TYPE ST_CamStatus :
STRUCT
    eState : E_CamMachineState;
    eProcessPhase : E_CamProcessPhase;
    bPowerEnabled : BOOL;
    bReferenced : BOOL;
    bRecipeLoaded : BOOL;
    bCamActive : BOOL;
    bRunning : BOOL;
    bBusy : BOOL;
    eApplicationError : E_CamApplicationError;
    eErrorSource : E_CamErrorSource;
    udiMotionErrorID : UDINT;
    lrCalculatedMaxSlaveVelocity : LREAL;
    lrCalculatedMaxSlaveAcceleration : LREAL;
    lrCalculatedMaxSlaveJerk : LREAL;
    lrCalculatedFaultStopSlaveAcceleration : LREAL;
    lrCalculatedFaultStopSlaveJerk : LREAL;
END_STRUCT
END_TYPE

(* stored: Version 1.1.0.1, ProductVersion 3.1.4024.16
   DUT ST_CamStatus: Id {fc009ade-7c77-4017-a2c5-fc4d406dae1c} *)
